Yaskawa INFORM job: 20211029ZUOGANGJIAOSAVE.JBI

/JOB
//NAME 20211029ZUOGANGJIAOSAVE
//POS
///NPOS 15,0,0,1,0,0
///TOOL 1
///POSTYPE PULSE
///PULSE
C00000=-6204,-15754,-18168,4454,-123898,-74311
C00001=-18321,-53773,-71210,-2327,-80039,-81868
C00002=-5575,-26998,-92017,-3234,-45195,-85018
C00003=-19625,-24229,-92072,-3290,-43470,-80509
C00004=-40364,-10263,-78411,-313,-44259,-47437
C00005=-32929,-5167,-69046,1265,-46694,-34744
C00006=-25417,20776,-43713,1030,-44670,-37067
C00007=-19212,27847,-31686,2815,-46500,-17389
C00008=-11867,28183,-27590,1845,-45132,5097
C00009=6393,26861,-34200,3324,-40364,1010
C00010=11035,23431,-36851,-2816,-38898,13574
C00011=20730,18312,-39742,-1088,-47602,36713
C00012=19793,13615,-53254,-1191,-41841,37081
C00013=34596,2740,-43617,410,-53764,32919
C00014=-1,-38943,-47654,0,-74515,0
///POSTYPE ROBOT
///RECTAN
///RCONF 0,0,0,0,0,0,0,0,0,0,0,0,0,0,0,0,0,0,0,0,0,0,0,0
P00001=629.883,8.042,-21.694,-154.9112,52.6025,29.7528
//INST
///DATE 2021/11/01 17:30
///ATTR SC,RW
///GROUP1 RB1
NOP
MOVJ C00000 VJ=10.00
MOVL C00001 V=20.0
MOVL C00002 V=20.0
CALL JOB:STARTDETPRG
WAIT B005=1
MOVL P001 V=23.0
CALL JOB:ENDDETPRG
CALL JOB:STARTCOR
ARCON AC=150 AV=25.0
MOVL C00003 V=20.0
CALL JOB:ENDDETPRG
ARCOF
MOVL C00004 V=20.0
MOVL C00005 V=20.0
CALL JOB:STARTDETPRG
WAIT B005=1
MOVL P001 V=23.0
CALL JOB:ENDDETPRG
CALL JOB:STARTCOR
ARCON AC=160 AV=25.0
MOVL C00006 V=20.0
CALL JOB:ENDDETPRG
ARCOF
MOVL C00007 V=20.0
MOVL C00008 V=20.0
CALL JOB:STARTDETPRG
WAIT B005=1
MOVL P001 V=23.0
CALL JOB:ENDDETPRG
CALL JOB:STARTCOR
ARCON AC=150 AV=25.0
MOVL C00009 V=20.0
CALL JOB:ENDDETPRG
ARCOF
MOVL C00010 V=20.0
MOVL C00011 V=20.0
CALL JOB:STARTDETPRG
WAIT B005=1
MOVL P001 V=23.0
CALL JOB:ENDDETPRG
CALL JOB:STARTCOR
ARCON AC=150 AV=25.0
MOVL C00012 V=20.0
CALL JOB:ENDDETPRG
ARCOF
MOVL C00013 V=20.0
MOVJ C00014 VJ=10.00
END
